Fanuc KAREL source: ka00109.KL

-- PROVISIONAL review KL for V940-1; original PC SHA256 558e20bca71038c82ebf4acb95377a896ff7e16cf1cc16cbb4e71fdd862c812a
-- Incomplete behavior may be omitted. Consult companion uncertainty JSON. Do not deploy.
PROGRAM KA00109
%NOLOCKGROUP
VAR
  DST : INTEGER
-- UNRESOLVED_DECL SRC type=00001c
BEGIN
  -- V9_ZERO_TABLE_METADATA_HINT layout=0001; no indexed target words; source/name/runtime held
  -- UNRESOLVED_PC offsets 5-15; opcodes 9D,22,A5
  -- UNRESOLVED_PC offsets 20-32; opcodes 21,23
  -- UNRESOLVED_PC offsets 37-41; opcodes 7F
END KA00109
